Fanuc KAREL source: kf00098.KL

-- PROVISIONAL review KL for V770-1; original PC SHA256 918c0b6de77b76153b5b829fade053a3103e54e1662064e3bc64cc1cc0f315b6
-- Incomplete behavior may be omitted. Consult companion uncertainty JSON. Do not deploy.
PROGRAM KF00098
%NOLOCKGROUP
BEGIN
  -- UNRESOLVED_PC offsets 5-16; opcodes 2E,23
  -- UNRESOLVED_PC offsets 21-32; opcodes 2E,23
  -- UNRESOLVED_PC offsets 37-55; opcodes 27,27,9D,22,22,31
  -- UNRESOLVED_PC offsets 60-64; opcodes 7F
END KF00098
